FUNCTION_BLOCK PID_CONTROLLER (* Whiteboard flag PID; direct atomic gain update; synthetic validation *)
  (* Standard: 61499-2 *)
  (* Version 0.1, 2026-10-18, Guilherme *)
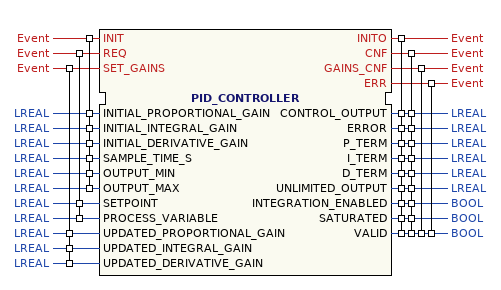
  EVENT_INPUT
    INIT WITH INITIAL_PROPORTIONAL_GAIN, INITIAL_INTEGRAL_GAIN, INITIAL_DERIVATIVE_GAIN, SAMPLE_TIME_S, OUTPUT_MIN, OUTPUT_MAX;
    REQ WITH SETPOINT, PROCESS_VARIABLE;
    SET_GAINS WITH UPDATED_PROPORTIONAL_GAIN, UPDATED_INTEGRAL_GAIN, UPDATED_DERIVATIVE_GAIN;
  END_EVENT
  EVENT_OUTPUT
    INITO WITH CONTROL_OUTPUT, ERROR, P_TERM, I_TERM, D_TERM, UNLIMITED_OUTPUT, INTEGRATION_ENABLED, SATURATED, VALID;
    CNF WITH CONTROL_OUTPUT, ERROR, P_TERM, I_TERM, D_TERM, UNLIMITED_OUTPUT, INTEGRATION_ENABLED, SATURATED, VALID;
    GAINS_CNF WITH VALID;
    ERR WITH VALID;
  END_EVENT
  VAR_INPUT
    INITIAL_PROPORTIONAL_GAIN : LREAL;
    INITIAL_INTEGRAL_GAIN : LREAL;
    INITIAL_DERIVATIVE_GAIN : LREAL;
    SAMPLE_TIME_S : LREAL;
    OUTPUT_MIN : LREAL;
    OUTPUT_MAX : LREAL;
    SETPOINT : LREAL;
    PROCESS_VARIABLE : LREAL;
    UPDATED_PROPORTIONAL_GAIN : LREAL;
    UPDATED_INTEGRAL_GAIN : LREAL;
    UPDATED_DERIVATIVE_GAIN : LREAL;
  END_VAR
  VAR_OUTPUT
    CONTROL_OUTPUT : LREAL;
    ERROR : LREAL;
    P_TERM : LREAL;
    I_TERM : LREAL;
    D_TERM : LREAL;
    UNLIMITED_OUTPUT : LREAL;
    INTEGRATION_ENABLED : BOOL;
    SATURATED : BOOL;
    VALID : BOOL;
  END_VAR
  VAR
    KP_ACTIVE : LREAL;
    KI_ACTIVE : LREAL;
    KD_ACTIVE : LREAL;
    TS_ACTIVE : LREAL;
    LOW : LREAL;
    HIGH : LREAL;
    I_MEMORY : LREAL;
    E_PREV : LREAL;
    E_NEXT : LREAL;
    I_NEXT : LREAL;
    D_NEXT : LREAL;
    P_NEXT : LREAL;
    IT_NEXT : LREAL;
    DT_NEXT : LREAL;
    RAW_NEXT : LREAL;
  END_VAR
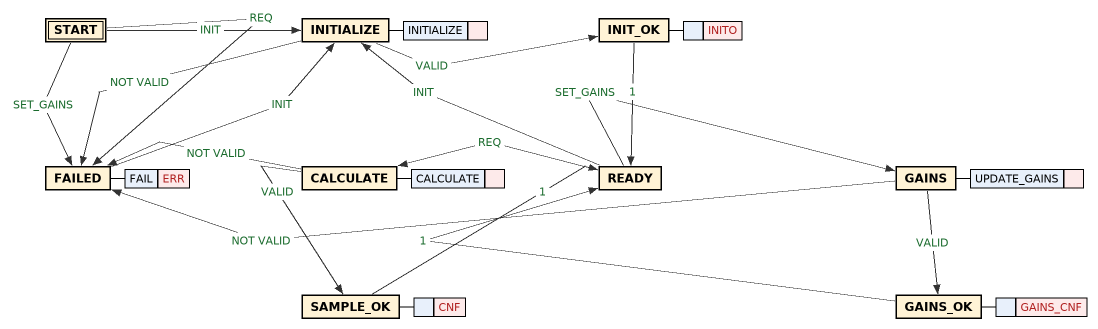
  EC_STATES
    START;
    INITIALIZE : INITIALIZE;
    INIT_OK : -> INITO;
    READY;
    CALCULATE : CALCULATE;
    SAMPLE_OK : -> CNF;
    GAINS : UPDATE_GAINS;
    GAINS_OK : -> GAINS_CNF;
    FAILED : FAIL -> ERR;
  END_STATES
  EC_TRANSITIONS
    START TO INITIALIZE := INIT;
    START TO FAILED := REQ;
    START TO FAILED := SET_GAINS;
    INITIALIZE TO INIT_OK := VALID;
    INITIALIZE TO FAILED := NOT VALID;
    INIT_OK TO READY := 1;
    READY TO INITIALIZE := INIT;
    READY TO GAINS := SET_GAINS;
    READY TO CALCULATE := REQ;
    CALCULATE TO SAMPLE_OK := VALID;
    CALCULATE TO FAILED := NOT VALID;
    SAMPLE_OK TO READY := 1;
    GAINS TO GAINS_OK := VALID;
    GAINS TO FAILED := NOT VALID;
    GAINS_OK TO READY := 1;
    FAILED TO INITIALIZE := INIT;
  END_TRANSITIONS
  ALGORITHM INITIALIZE IN ST:
VALID := (INITIAL_PROPORTIONAL_GAIN >= -1.0E+100) AND (INITIAL_PROPORTIONAL_GAIN <= 1.0E+100) AND (INITIAL_INTEGRAL_GAIN >= -1.0E+100) AND (INITIAL_INTEGRAL_GAIN <= 1.0E+100) AND (INITIAL_DERIVATIVE_GAIN >= -1.0E+100) AND (INITIAL_DERIVATIVE_GAIN <= 1.0E+100) AND (SAMPLE_TIME_S >= -1.0E+100) AND (SAMPLE_TIME_S <= 1.0E+100) AND (OUTPUT_MIN >= -1.0E+100) AND (OUTPUT_MIN <= 1.0E+100) AND (OUTPUT_MAX >= -1.0E+100) AND (OUTPUT_MAX <= 1.0E+100) AND (SAMPLE_TIME_S > 0.0) AND (OUTPUT_MIN < OUTPUT_MAX);
IF VALID THEN
    KP_ACTIVE := INITIAL_PROPORTIONAL_GAIN;
    KI_ACTIVE := INITIAL_INTEGRAL_GAIN;
    KD_ACTIVE := INITIAL_DERIVATIVE_GAIN;
    TS_ACTIVE := SAMPLE_TIME_S;
    LOW := OUTPUT_MIN;
    HIGH := OUTPUT_MAX;
    I_MEMORY := 0.0;
    E_PREV := 0.0;
    INTEGRATION_ENABLED := TRUE;
    CONTROL_OUTPUT := 0.0;
    UNLIMITED_OUTPUT := 0.0;
    ERROR := 0.0;
    P_TERM := 0.0;
    I_TERM := 0.0;
    D_TERM := 0.0;
    SATURATED := FALSE;
END_IF;
  END_ALGORITHM
  ALGORITHM CALCULATE IN ST:
VALID := (SETPOINT >= -1.0E+100) AND (SETPOINT <= 1.0E+100) AND (PROCESS_VARIABLE >= -1.0E+100) AND (PROCESS_VARIABLE <= 1.0E+100);
IF VALID THEN
    E_NEXT := SETPOINT - PROCESS_VARIABLE;
    I_NEXT := I_MEMORY;
    IF INTEGRATION_ENABLED THEN
        I_NEXT := I_MEMORY + (TS_ACTIVE / 2.0) * (E_NEXT + E_PREV);
    END_IF;
    D_NEXT := (E_NEXT - E_PREV) / TS_ACTIVE;
    P_NEXT := KP_ACTIVE * E_NEXT;
    IT_NEXT := KI_ACTIVE * I_NEXT;
    DT_NEXT := KD_ACTIVE * D_NEXT;
    RAW_NEXT := P_NEXT + IT_NEXT + DT_NEXT;
    VALID := (E_NEXT >= -1.0E+100) AND (E_NEXT <= 1.0E+100) AND (I_NEXT >= -1.0E+100) AND (I_NEXT <= 1.0E+100) AND (D_NEXT >= -1.0E+100) AND (D_NEXT <= 1.0E+100) AND (P_NEXT >= -1.0E+100) AND (P_NEXT <= 1.0E+100) AND (IT_NEXT >= -1.0E+100) AND (IT_NEXT <= 1.0E+100) AND (DT_NEXT >= -1.0E+100) AND (DT_NEXT <= 1.0E+100) AND (RAW_NEXT >= -1.0E+100) AND (RAW_NEXT <= 1.0E+100);
    IF VALID THEN
        CONTROL_OUTPUT := RAW_NEXT;
        INTEGRATION_ENABLED := TRUE;
        SATURATED := FALSE;
        IF RAW_NEXT > HIGH THEN
            CONTROL_OUTPUT := HIGH;
            INTEGRATION_ENABLED := FALSE;
            SATURATED := TRUE;
        END_IF;
        IF RAW_NEXT < LOW THEN
            CONTROL_OUTPUT := LOW;
            INTEGRATION_ENABLED := FALSE;
            SATURATED := TRUE;
        END_IF;
        I_MEMORY := I_NEXT;
        E_PREV := E_NEXT;
        ERROR := E_NEXT;
        P_TERM := P_NEXT;
        I_TERM := IT_NEXT;
        D_TERM := DT_NEXT;
        UNLIMITED_OUTPUT := RAW_NEXT;
    END_IF;
END_IF;
  END_ALGORITHM
  ALGORITHM UPDATE_GAINS IN ST:
VALID := (UPDATED_PROPORTIONAL_GAIN >= -1.0E+100) AND (UPDATED_PROPORTIONAL_GAIN <= 1.0E+100) AND (UPDATED_INTEGRAL_GAIN >= -1.0E+100) AND (UPDATED_INTEGRAL_GAIN <= 1.0E+100) AND (UPDATED_DERIVATIVE_GAIN >= -1.0E+100) AND (UPDATED_DERIVATIVE_GAIN <= 1.0E+100);
IF VALID THEN
    KP_ACTIVE := UPDATED_PROPORTIONAL_GAIN;
    KI_ACTIVE := UPDATED_INTEGRAL_GAIN;
    KD_ACTIVE := UPDATED_DERIVATIVE_GAIN;
END_IF;
  END_ALGORITHM
  ALGORITHM FAIL IN ST:
VALID := FALSE;
  END_ALGORITHM
END_FUNCTION_BLOCK
